# EPICS substitutions: db/Beckhoff_5XXX/ecmcEL5101.substitutions
file "ecmcEL5101-chX.template"
{
    pattern {CH_ID}
            {01   }

}
